{attribute 'linkalways'} 
{attribute 'no_explicit_call' := 'This FB is a CLASS and must be accessed using methods or properties'}
{attribute 'enable_dynamic_creation'}
FUNCTION_BLOCK _Array0to2OfUSINT EXTENDS ArrayDatatypeBase_1D
VAR CONSTANT
	lBound : DINT := 0;
	uBound : DINT := 2;
END_VAR
VAR
	localData : ARRAY [lBound..uBound] OF USINT;
	activeData : REFERENCE TO ARRAY [lBound..uBound] OF USINT REF= localData;
	elements : ARRAY [lBound..uBound] OF _USINT(0);
	baseType : _USINT(0);
END_VAR

PROPERTY PUBLIC Address : PVOID
GET
Address := ADR(activeData);
END_GET
END_PROPERTY

PROPERTY PUBLIC BaseDatatype : I_Datatype
GET
BaseDatatype := baseType;
END_GET
END_PROPERTY

METHOD PUBLIC ClearReference
VAR_INPUT
END_VAR
activeData REF= localData;
SetElementReference();
END_METHOD

METHOD PUBLIC Clone : I_Datatype
VAR
    pClone : POINTER TO _Array0to2OfUSINT;
END_VAR
pClone := __NEW(_Array0to2OfUSINT());
pClone^.Value := Value;
Clone := pClone^;
END_METHOD

METHOD FB_init : BOOL
VAR_INPUT
	bInitRetains : BOOL; // if TRUE, the retain variables are initialized (warm start / cold start)
	bInCopyCode : BOOL;  // if TRUE, the instance afterwards gets moved into the copy code (online change)
END_VAR
SetElementReference();
END_METHOD

METHOD PUBLIC MakeReferenceTo
VAR_INPUT
	ReferenceTarget : REFERENCE TO ARRAY [lBound..uBound] OF USINT;
END_VAR
activeData REF= ReferenceTarget;
SetElementReference();
END_METHOD

METHOD PROTECTED OnSerializeArrayValues
VAR_INPUT
	Serializer : I_Serializer;
END_VAR
VAR
	i : DINT;
END_VAR
FOR i := lBound TO uBound DO
	elements[i].SerializeWith(Serializer);
END_FOR
END_METHOD

METHOD PROTECTED SetElementReference
VAR_INPUT
END_VAR
VAR
	i : DINT;
END_VAR
FOR i := lBound TO uBound DO
	elements[i].MakeReferenceTo(activeData[i]);
END_FOR
END_METHOD

PROPERTY PUBLIC Size : UDINT
GET
Size := SIZEOF(activeData);
END_GET
END_PROPERTY

METHOD PROTECTED TryDeserializeArrayValues : BOOL
VAR_INPUT
	Deserializer : I_Deserializer;
	Feedback : I_DeserializerFeedback;
END_VAR
VAR
	failed : BOOL;
	enumerator : I_DeserializerArrayForwardEnumerator;
	i : DINT;
END_VAR
enumerator := Deserializer.GetArrayEnumerator();
i := lBound;

WHILE enumerator.MoveNext() AND i <= uBound AND NOT failed DO
	
	IF NOT elements[i].TryDeserializeFrom(enumerator.Current, Feedback) THEN
		failed := TRUE;
		EXIT;
	END_IF
	i := i + 1;

END_WHILE
enumerator.Dispose();

TryDeserializeArrayValues := NOT failed;
END_METHOD

METHOD PUBLIC TryGetElementAsDatatypeByIndex : BOOL
VAR_INPUT
	Index : DINT;
	Destination : REFERENCE TO I_Datatype;
END_VAR
IF Index < lbound OR Index > ubound THEN
	RETURN;
END_IF

Destination := elements[Index];
TryGetElementAsDatatypeByIndex := TRUE;
END_METHOD

METHOD PUBLIC TryGetLowerBound : BOOL
VAR_INPUT
	Dimention : UDINT;
	Destination : REFERENCE TO DINT;
END_VAR
IF Dimention = 1 THEN
	Destination := lBound;
	TryGetLowerBound := TRUE;
END_IF
END_METHOD

METHOD PUBLIC TryGetUpperBound : BOOL
VAR_INPUT
	Dimention : UDINT;
	Destination : REFERENCE TO DINT;
END_VAR
IF Dimention = 1 THEN
	Destination := uBound;
	TryGetUpperBound := TRUE;
END_IF
END_METHOD

METHOD TryMakeReferenceTo : BOOL
VAR_INPUT
	Target : I_Datatype;
END_VAR
VAR
	pTargetData : POINTER TO ARRAY [lBound..uBound] OF USINT;
END_VAR
IF NOT IsEquivalentTo(Target) THEN
	RETURN;
END_IF

pTargetData := Target.Address;
activeData REF= pTargetData^;
SetElementReference();
TryMakeReferenceTo := TRUE;
END_METHOD

PROPERTY PUBLIC Value : REFERENCE TO ARRAY [lBound..uBound] OF USINT;
GET
Value ref= activeData;
END_GET
END_PROPERTY

END_FUNCTION_BLOCK

(* stored: Version 1.1.0.1, ProductVersion 3.1.4024.13
   POU _Array0to2OfUSINT: Id {97ba6251-0797-08ad-20c4-a811d2a463cd}, SpecialFunc None
   Folder Core: Id {d40f1a96-b607-0308-1a4d-91811eb1f640}
   Folder Constructor: Id {27a99c7c-f8b4-0b23-02e7-9a9be14c970d}
   Folder Protected: Id {b5dd3a28-8147-093f-1ac4-9c3e80e8b715}
   Folder Customize: Id {0b04ff73-2076-0098-3463-8f276c6c7a5a}
   Property Address: Id {7c7efdf8-17ae-008f-0226-4930925424e7}
   Get Get: Id {cb91481a-070a-0343-3c7c-c7ad10fb8d84}
   Property BaseDatatype: Id {6564742d-9082-095b-15c6-623c3ac7c6de}
   Get Get: Id {3dc79983-8c2f-01ed-1906-ff642c4f4598}
   Method ClearReference: Id {24191594-fb34-0855-2bce-a922995581d7}
   Method Clone: Id {78cdaf05-3d2f-0d2e-1878-6b9e44e5057d}
   Method FB_init: Id {5da9a1fe-c111-0f20-23d8-168b6e42e286}
   Method MakeReferenceTo: Id {3c225855-8ae7-0149-3ecf-9e8a1a5ab443}
   Method OnSerializeArrayValues: Id {3300385d-c4eb-0da8-0132-53fb85ff7e6d}
   Method SetElementReference: Id {38e4ac71-6436-0376-362a-271f360fe578}
   Property Size: Id {06ffd24a-c7a0-0160-38a7-8fc5849e597c}
   Get Get: Id {e7f03b69-a0e8-05b0-0a41-63b1c12f0379}
   Method TryDeserializeArrayValues: Id {f3e39256-012e-0882-0e51-133b4d5ce1dd}
   Method TryGetElementAsDatatypeByIndex: Id {46aed853-f5a6-05dc-3d64-f290d4e5c60c}
   Method TryGetLowerBound: Id {cb7014f3-1ae4-02aa-20a3-a862b1c7d8f7}
   Method TryGetUpperBound: Id {25518b62-0495-0327-1887-6639da74981a}
   Method TryMakeReferenceTo: Id {b3a722ae-c8ae-0410-26b5-ca5c2e4fd661}
   Property Value: Id {0b3cb14b-e52a-0865-0a82-426d566d3bd0}
   Get Get: Id {9695706b-6b33-0379-3cc2-86199b0683b0} *)
